(* IEC 61131-3 sources: plc-iiot-stack/src/POUs/Iiot/FB_MqttCommands, 19 files *)

(* ---- FB_MqttCommands.decl.st ---- *)
// Назначение: шлюз команд MQTT (data_schema 5): подписка <prefix>/+/cmd/+ (QoS 1), разбор подмножества JSON,
//             проверки по порядку раздела 5.1 (retained, invalid_payload, unsupported_version, topic_mismatch,
//             not_whitelisted, out_of_range, expired, duplicate, rate_limited) и ответ в
//             <prefix>/<device>/cmd_ack/<command>. Сообщение не своей станции или без читаемого cmd_id —
//             без ответа (udiDropped). Прошедшая команда — импульс xCmdValid и stCmd: вызывающий пишет её в
//             GVL_Hmi и вызывает Arm(); дальше ФБ ждёт, пока устройство увеличит uiCmdSeq (ok или
//             device_rejected по eCmdResult), иначе через tDeviceTimeout — timeout. Значения (SpeedSp) ФБ
//             устройства не квитирует: ok — сразу после записи. Одна команда в обработке за раз.
// Автор:      kr0nsch
// Версия:     0.1.0
// Документ:   docs/plc_mqtt.md, раздел «Команды»
FUNCTION_BLOCK FB_MqttCommands
VAR_INPUT
    xEnable : BOOL;
    itfClient : I_MqttClient;
    ltNow : LTIME;                                            // монотонное время (LTIME())
    uliTs_ms : ULINT;                                         // время UTC, мс: проверка ts и поле ts ответа
    sTopicPrefix : STRING(GVL_Const.IIOT_PREFIX_LEN);         // site/area/unit
    uiDevSeq : UINT;                                          // uiCmdSeq устройства команды в обработке
    iDevResult : INT;                                         // eCmdResult того же устройства
    tMaxAge : TIME := GVL_Const.CMD_MAX_AGE;
    tDeviceTimeout : TIME := GVL_Const.CMD_DEVICE_TIMEOUT;
    uiRateLimit : UINT := GVL_Const.CMD_RATE_LIMIT;           // не больше CMD_RATE_LIMIT
    tRateWindow : TIME := GVL_Const.CMD_RATE_WINDOW;
    uiMaxPerCycle : UINT := GVL_Const.CMD_MAX_PER_CYCLE;
END_VAR
VAR_IN_OUT
    aRules : ARRAY[*] OF ST_IiotCmdRule;                      // белый список
END_VAR
VAR_OUTPUT
    xCmdValid : BOOL;                                         // в этом вызове: записать stCmd в GVL_Hmi, затем Arm()
    stCmd : ST_IiotCmd;
    xPending : BOOL;                                          // ждём обработки устройством
    xSubscribed : BOOL;
    eLastReason : E_IiotCmdReason := E_IiotCmdReason.Ok;
    udiReceived : UDINT;
    udiAccepted : UDINT;                                      // ответов ok
    udiRejected : UDINT;                                      // ответов с отказом
    udiDropped : UDINT;                                       // без ответа: чужой топик, нет cmd_id
    udiAckFailed : UDINT;                                     // ответ не принят клиентом или не помещается
END_VAR
VAR
    fbParser : FB_JsonFlatParser;
    fbJson : FB_JsonBuilder;
    sFilter : STRING(GVL_Const.MQTT_TOPIC_LEN);
    sRxTopic : STRING(GVL_Const.MQTT_TOPIC_LEN);
    sRxPayload : STRING(GVL_Const.MQTT_CMD_PAYLOAD_LEN);
    xRxTruncated : BOOL;
    xRxRetained : BOOL;
    sAckTopic : STRING(GVL_Const.MQTT_TOPIC_LEN);
    // команда, на которую готовится ответ
    sTopicDevice : STRING(GVL_Const.IIOT_LEVEL_LEN);
    sTopicCommand : STRING(GVL_Const.IIOT_LEVEL_LEN);
    sCmdId : STRING(GVL_Const.JSON_STR_LEN);
    // повторы и частота
    aHistory : ARRAY[1..GVL_Const.CMD_HISTORY_LEN] OF STRING(GVL_Const.CMD_ID_LEN);
    uiHistoryNext : UINT := 1;
    aRateTimes : ARRAY[1..GVL_Const.CMD_RATE_LIMIT] OF LTIME;   // моменты последних прошедших команд
    uiRateNext : UINT := 1;
    uiRateCount : UINT;
    // обработка устройством
    xAwaitArm : BOOL;
    uiSeqArmed : UINT;
    ltPendingSince : LTIME;
    uiMsg : UINT;
END_VAR

(* ---- Arm.method.decl.st ---- *)
// Вызвать после записи stCmd в GVL_Hmi в том же цикле: uiSeqBefore — uiCmdSeq устройства до записи.
// Команды-значения (SpeedSp, SubstValue) отвечают ok сразу: ФБ устройства их не квитирует.
METHOD Arm
VAR_INPUT
    uiSeqBefore : UINT;
END_VAR

(* ---- Arm.method.impl.st ---- *)
IF NOT xAwaitArm THEN
    RETURN;
END_IF
xAwaitArm := FALSE;
IF F_IiotCmdKind(eCommand := stCmd.eCommand) = E_IiotCmdKind.Value THEN
    Finish(eReason := E_IiotCmdReason.Ok, iCmdResult := 0);
ELSE
    uiSeqArmed := uiSeqBefore;
    ltPendingSince := ltNow;
    xPending := TRUE;
END_IF

(* ---- Check.method.decl.st ---- *)
// Проверки шлюза по порядку data_schema 5.1, пункты 1–9; Ok — stCmd заполнена, момент учтён в частоте.
METHOD PRIVATE Check : E_IiotCmdReason
VAR_IN_OUT
    aRuleTable : ARRAY[*] OF ST_IiotCmdRule;
END_VAR
VAR
    sText : STRING(GVL_Const.JSON_STR_LEN);
    sKey : STRING(GVL_Const.JSON_KEY_LEN);
    iMajor : INT;
    uiIdx : UINT;
    lrTs : LREAL;
    lrValue : LREAL;
    lrMin : LREAL;
    lrMax : LREAL;
    xHasValue : BOOL;
    eCommand : E_IiotCommand;
    eKind : E_IiotCmdKind;
    diRule : DINT;
END_VAR

(* ---- Check.method.impl.st ---- *)
// 1. retained
IF xRxRetained THEN
    Check := E_IiotCmdReason.Retained;
    RETURN;
END_IF
// 2. состав и типы полей (command.schema.json; диапазон value — в п. 6)
Check := E_IiotCmdReason.InvalidPayload;
IF NOT fbParser.GetString(sKey := 'schema_version', sValue := sText) THEN
    RETURN;
END_IF
iMajor := F_IiotSchemaMajor(sVersion := sText);
IF iMajor < 0 THEN
    RETURN;
END_IF
FOR uiIdx := 1 TO fbParser.uiCount DO
    sKey := fbParser.KeyAt(uiIdx := uiIdx);
    IF sKey <> 'schema_version' AND sKey <> 'cmd_id' AND sKey <> 'ts' AND sKey <> 'origin' AND sKey <> 'command'
       AND sKey <> 'value' THEN
        RETURN;                     // лишнее поле: схема команды строгая
    END_IF
END_FOR
IF NOT fbParser.FieldIsInteger(sKey := 'ts') OR NOT fbParser.GetNumber(sKey := 'ts', lrValue := lrTs) THEN
    RETURN;
END_IF
IF lrTs < ULINT_TO_LREAL(GVL_Const.TS_MIN_MS) OR lrTs > ULINT_TO_LREAL(GVL_Const.TS_MAX_MS) THEN
    RETURN;
END_IF
IF NOT fbParser.GetString(sKey := 'origin', sValue := sText) THEN
    RETURN;
END_IF
IF NOT F_IiotIsPrintable(sText := sText, iMaxLen := UINT_TO_INT(GVL_Const.CMD_ORIGIN_LEN)) THEN
    RETURN;
END_IF
IF NOT fbParser.GetString(sKey := 'command', sValue := sText) THEN
    RETURN;
END_IF
eCommand := F_IiotCmdFromString(sCommand := sText);
IF eCommand = E_IiotCommand.None THEN
    RETURN;
END_IF
eKind := F_IiotCmdKind(eCommand := eCommand);
xHasValue := fbParser.FieldType(sKey := 'value') <> E_JsonType.Missing;
IF xHasValue AND NOT fbParser.GetNumber(sKey := 'value', lrValue := lrValue) THEN
    RETURN;                         // value не число
END_IF
IF eKind = E_IiotCmdKind.Pulse AND xHasValue THEN
    RETURN;                         // value у импульсной команды
END_IF
IF eKind <> E_IiotCmdKind.Pulse AND NOT xHasValue THEN
    RETURN;                         // нет value
END_IF
IF eKind = E_IiotCmdKind.Mask
   AND (NOT fbParser.FieldIsInteger(sKey := 'value') OR lrValue < 0.0 OR lrValue > GVL_Const.CMD_MASK_MAX) THEN
    RETURN;                         // маска: целое 0..65535
END_IF
// 3. мажорная версия
IF iMajor <> UINT_TO_INT(GVL_Const.IIOT_SCHEMA_MAJOR) THEN
    Check := E_IiotCmdReason.UnsupportedVersion;
    RETURN;
END_IF
// 4. команда в теле и в топике
IF sText <> sTopicCommand THEN
    Check := E_IiotCmdReason.TopicMismatch;
    RETURN;
END_IF
// 5. белый список
diRule := FindRule(aRuleTable := aRuleTable, eCommandIn := eCommand);
IF diRule < LOWER_BOUND(aRuleTable, 1) THEN
    Check := E_IiotCmdReason.NotWhitelisted;
    RETURN;
END_IF
// 6. диапазон значения
IF xHasValue THEN
    IF aRuleTable[diRule].xRange THEN
        lrMin := REAL_TO_LREAL(aRuleTable[diRule].rMin);
        lrMax := REAL_TO_LREAL(aRuleTable[diRule].rMax);
    ELSE
        lrMin := -GVL_Const.REAL_ABS_MAX;
        lrMax := GVL_Const.REAL_ABS_MAX;
    END_IF
    IF eCommand = E_IiotCommand.SpeedSp THEN       // схема: 0..100 % независимо от белого списка
        lrMin := MAX(lrMin, GVL_Const.SPEED_SP_MIN_PCT);
        lrMax := MIN(lrMax, GVL_Const.SPEED_SP_MAX_PCT);
    END_IF
    IF lrValue < lrMin OR lrValue > lrMax THEN
        Check := E_IiotCmdReason.OutOfRange;
        RETURN;
    END_IF
END_IF
// 7. возраст ts (часы ПЛК должны быть установлены)
IF NOT F_IiotClockValid(uliTs_ms := uliTs_ms)
   OR ABS(ULINT_TO_LREAL(uliTs_ms) - lrTs) > ULINT_TO_LREAL(TIME_TO_ULINT(tMaxAge)) THEN
    Check := E_IiotCmdReason.Expired;
    RETURN;
END_IF
// 8. повтор cmd_id
IF IsDuplicate() THEN
    Check := E_IiotCmdReason.Duplicate;
    RETURN;
END_IF
// 9. частота
IF NOT RateAllows() THEN
    Check := E_IiotCmdReason.RateLimited;
    RETURN;
END_IF
stCmd.diRule := diRule;
stCmd.sDevice := sTopicDevice;
stCmd.sCommand := sTopicCommand;
stCmd.eCommand := eCommand;
stCmd.rValue := LREAL_TO_REAL(lrValue);
stCmd.sCmdId := sCmdId;
Check := E_IiotCmdReason.Ok;

(* ---- FB_MqttCommands.impl.st ---- *)
xCmdValid := FALSE;
IF NOT xEnable OR itfClient = 0 THEN
    xSubscribed := FALSE;
    xPending := FALSE;
    xAwaitArm := FALSE;
    RETURN;
END_IF
IF NOT itfClient.IsConnected() THEN
    xSubscribed := FALSE;     // после подключения — подписка заново (сессия может быть чистой)
    RETURN;
END_IF
IF NOT xSubscribed THEN
    sFilter := CONCAT(sTopicPrefix, GVL_Const.TOPIC_CMD_FILTER_SUFFIX);
    xSubscribed := itfClient.Subscribe(sTopicFilter := sFilter, eQos := E_MqttQos.AtLeastOnce);
    IF NOT xSubscribed THEN
        RETURN;
    END_IF
END_IF

// Команда прошла проверки в прошлом вызове, но Arm() не вызван: до устройства она не дошла
IF xAwaitArm THEN
    xAwaitArm := FALSE;
    Finish(eReason := E_IiotCmdReason.Timeout, iCmdResult := 0);
END_IF
// Команда в обработке устройством
IF xPending THEN
    IF uiDevSeq <> uiSeqArmed AND iDevResult >= GVL_Const.CMD_RESULT_ACCEPTED
       AND iDevResult <= GVL_Const.CMD_RESULT_LAST THEN
        xPending := FALSE;
        IF iDevResult = GVL_Const.CMD_RESULT_ACCEPTED THEN
            Finish(eReason := E_IiotCmdReason.Ok, iCmdResult := iDevResult);
        ELSE
            Finish(eReason := E_IiotCmdReason.DeviceRejected, iCmdResult := iDevResult);
        END_IF
    ELSIF ltNow < ltPendingSince THEN
        ltPendingSince := ltNow;
    ELSIF (ltNow - ltPendingSince) >= TIME_TO_LTIME(tDeviceTimeout) THEN
        xPending := FALSE;
        Finish(eReason := E_IiotCmdReason.Timeout, iCmdResult := 0);
    END_IF
    IF xPending THEN
        RETURN;
    END_IF
END_IF

FOR uiMsg := 1 TO MAX(uiMaxPerCycle, 1) DO
    IF xCmdValid THEN
        EXIT;
    END_IF
    IF NOT itfClient.Receive(sTopic := sRxTopic, sPayload := sRxPayload, xTruncated => xRxTruncated,
                             xRetained => xRxRetained) THEN
        EXIT;
    END_IF
    udiReceived := udiReceived + 1;
    HandleMessage(aRuleTable := aRules);
END_FOR

(* ---- FindRule.method.decl.st ---- *)
// Строка белого списка для (sTopicDevice, eCommandIn); нет — LOWER_BOUND - 1.
METHOD PRIVATE FindRule : DINT
VAR_IN_OUT
    aRuleTable : ARRAY[*] OF ST_IiotCmdRule;
END_VAR
VAR_INPUT
    eCommandIn : E_IiotCommand;
END_VAR
VAR
    diIdx : DINT;
END_VAR

(* ---- FindRule.method.impl.st ---- *)
FindRule := LOWER_BOUND(aRuleTable, 1) - 1;
FOR diIdx := LOWER_BOUND(aRuleTable, 1) TO UPPER_BOUND(aRuleTable, 1) DO
    IF aRuleTable[diIdx].eCommand = eCommandIn AND aRuleTable[diIdx].sDevice = sTopicDevice THEN
        FindRule := diIdx;
        RETURN;
    END_IF
END_FOR

(* ---- Finish.method.decl.st ---- *)
// Ответ в <prefix>/<sTopicDevice>/cmd_ack/<sTopicCommand>: schema_version, cmd_id, ts, command, result, reason
// и cmd_result (device_rejected). Счётчики принятых и отклонённых команд.
METHOD PRIVATE Finish
VAR_INPUT
    eReason : E_IiotCmdReason;
    iCmdResult : INT;             // E_CmdResult устройства; 0 — нет
END_VAR
VAR
    sResultText : STRING(GVL_Const.IIOT_TEXT_LEN);
    sPath : STRING(GVL_Const.MQTT_TOPIC_LEN);
END_VAR

(* ---- Finish.method.impl.st ---- *)
eLastReason := eReason;
IF eReason = E_IiotCmdReason.Ok THEN
    udiAccepted := udiAccepted + 1;
ELSE
    udiRejected := udiRejected + 1;
END_IF
sPath := CONCAT(CONCAT(sTopicDevice, GVL_Const.TOPIC_SEPARATOR), GVL_Const.TOPIC_ACK_LEVEL);
sPath := CONCAT(CONCAT(sPath, GVL_Const.TOPIC_SEPARATOR), sTopicCommand);
sAckTopic := F_IiotTopic(sPrefix := sTopicPrefix, sPath := sPath);
fbJson.Begin();
fbJson.AddString(sKey := 'schema_version', sValue := GVL_Const.IIOT_SCHEMA_VERSION);
fbJson.AddString(sKey := 'cmd_id', sValue := sCmdId);
fbJson.AddInt(sKey := 'ts', liValue := ULINT_TO_LINT(uliTs_ms));
fbJson.AddString(sKey := 'command', sValue := sTopicCommand);
IF eReason = E_IiotCmdReason.Ok THEN
    fbJson.AddString(sKey := 'result', sValue := 'accepted');
ELSE
    fbJson.AddString(sKey := 'result', sValue := 'rejected');
END_IF
fbJson.AddString(sKey := 'reason', sValue := F_IiotCmdReasonText(eReason := eReason));
sResultText := F_IiotCmdResultText(iResult := iCmdResult);
IF eReason = E_IiotCmdReason.DeviceRejected AND LEN(sResultText) > 0 THEN
    fbJson.AddString(sKey := 'cmd_result', sValue := sResultText);
END_IF
IF NOT fbJson.Finish() OR LEN(sAckTopic) = 0 THEN
    udiAckFailed := udiAckFailed + 1;
ELSIF NOT itfClient.Publish(sTopic := sAckTopic, eQos := E_MqttQos.AtLeastOnce, xRetain := FALSE,
                            sPayload := fbJson.sJson) THEN
    udiAckFailed := udiAckFailed + 1;
END_IF

(* ---- HandleMessage.method.decl.st ---- *)
// Разбор принятого сообщения: без ответа (чужой топик, нет cmd_id), отказ с ответом или команда в stCmd.
METHOD PRIVATE HandleMessage
VAR_IN_OUT
    aRuleTable : ARRAY[*] OF ST_IiotCmdRule;
END_VAR
VAR
    eReason : E_IiotCmdReason;
END_VAR

(* ---- HandleMessage.method.impl.st ---- *)
sCmdId := '';
IF NOT SplitTopic() THEN
    udiDropped := udiDropped + 1;      // не команда своей станции — отвечать некуда
    RETURN;
END_IF
IF xRxTruncated OR NOT fbParser.Parse(sJson := sRxPayload) THEN
    udiDropped := udiDropped + 1;      // не JSON-объект: cmd_id не прочитать
    RETURN;
END_IF
IF NOT fbParser.GetString(sKey := 'cmd_id', sValue := sCmdId) OR NOT F_IiotIsCmdId(sText := sCmdId) THEN
    sCmdId := '';
    udiDropped := udiDropped + 1;
    RETURN;
END_IF
eReason := Check(aRuleTable := aRuleTable);
IF eReason <> E_IiotCmdReason.Duplicate THEN
    Remember();
END_IF
IF eReason = E_IiotCmdReason.Ok THEN
    xCmdValid := TRUE;
    xAwaitArm := TRUE;
ELSE
    Finish(eReason := eReason, iCmdResult := 0);
END_IF

(* ---- IsDuplicate.method.decl.st ---- *)
// cmd_id текущей команды встречался среди последних CMD_HISTORY_LEN.
METHOD PRIVATE IsDuplicate : BOOL
VAR
    uiIdx : UINT;
END_VAR

(* ---- IsDuplicate.method.impl.st ---- *)
FOR uiIdx := 1 TO GVL_Const.CMD_HISTORY_LEN DO
    IF LEN(aHistory[uiIdx]) > 0 AND aHistory[uiIdx] = sCmdId THEN
        IsDuplicate := TRUE;
        RETURN;
    END_IF
END_FOR

(* ---- RateAllows.method.decl.st ---- *)
// Частота: не больше uiRateLimit прошедших команд за tRateWindow. TRUE — команда разрешена и учтена.
METHOD PRIVATE RateAllows : BOOL
VAR
    uiLimit : UINT;
END_VAR

(* ---- RateAllows.method.impl.st ---- *)
uiLimit := MIN(MAX(uiRateLimit, 1), GVL_Const.CMD_RATE_LIMIT);
IF uiRateNext < 1 OR uiRateNext > uiLimit THEN
    uiRateNext := 1;
END_IF
// в кольце из uiLimit моментов следующая позиция — самая старая из последних uiLimit команд
IF uiRateCount >= uiLimit AND_THEN ltNow >= aRateTimes[uiRateNext]
   AND_THEN (ltNow - aRateTimes[uiRateNext]) <= TIME_TO_LTIME(tRateWindow) THEN
    RETURN;
END_IF
aRateTimes[uiRateNext] := ltNow;
uiRateNext := uiRateNext + 1;
IF uiRateNext > uiLimit THEN
    uiRateNext := 1;
END_IF
IF uiRateCount < uiLimit THEN
    uiRateCount := uiRateCount + 1;
END_IF
RateAllows := TRUE;

(* ---- Remember.method.impl.st ---- *)
IF uiHistoryNext < 1 OR uiHistoryNext > GVL_Const.CMD_HISTORY_LEN THEN
    uiHistoryNext := 1;
END_IF
aHistory[uiHistoryNext] := sCmdId;
uiHistoryNext := uiHistoryNext + 1;

(* ---- SplitTopic.method.decl.st ---- *)
// Разобрать sRxTopic вида <prefix>/<DEVICE>/cmd/<Command> в sTopicDevice и sTopicCommand. FALSE — топик не
// своей станции или уровни не по шаблонам ([A-Z][A-Z0-9_]{0,15} и [A-Za-z][A-Za-z0-9_]{0,31}).
METHOD PRIVATE SplitTopic : BOOL
VAR
    iPrefixLen : INT;
    sRest : STRING(GVL_Const.MQTT_TOPIC_LEN);
    sTail : STRING(GVL_Const.MQTT_TOPIC_LEN);
    iSlash : INT;
END_VAR

(* ---- SplitTopic.method.impl.st ---- *)
sTopicDevice := '';
sTopicCommand := '';
iPrefixLen := LEN(sTopicPrefix);
IF iPrefixLen = 0 OR LEN(sRxTopic) <= iPrefixLen + 1 THEN
    RETURN;
END_IF
IF LEFT(sRxTopic, iPrefixLen) <> sTopicPrefix OR MID(sRxTopic, 1, iPrefixLen + 1) <> GVL_Const.TOPIC_SEPARATOR THEN
    RETURN;
END_IF
sRest := RIGHT(sRxTopic, LEN(sRxTopic) - iPrefixLen - 1);
// <DEVICE>
iSlash := FIND(sRest, GVL_Const.TOPIC_SEPARATOR);
IF iSlash <= 1 OR iSlash - 1 > UINT_TO_INT(GVL_Const.IIOT_DEVICE_LEN) THEN
    RETURN;
END_IF
sTopicDevice := LEFT(sRest, iSlash - 1);
sTail := RIGHT(sRest, LEN(sRest) - iSlash);
// cmd
iSlash := FIND(sTail, GVL_Const.TOPIC_SEPARATOR);
IF iSlash <= 1 OR LEFT(sTail, iSlash - 1) <> GVL_Const.TOPIC_CMD_LEVEL THEN
    sTopicDevice := '';
    RETURN;
END_IF
// <Command>
IF LEN(sTail) - iSlash > UINT_TO_INT(GVL_Const.IIOT_LEVEL_LEN) THEN
    sTopicDevice := '';
    RETURN;
END_IF
sTopicCommand := RIGHT(sTail, LEN(sTail) - iSlash);
IF NOT F_IiotIsName(sText := sTopicDevice, iMaxLen := UINT_TO_INT(GVL_Const.IIOT_DEVICE_LEN), xUpperOnly := TRUE)
   OR NOT F_IiotIsName(sText := sTopicCommand, iMaxLen := UINT_TO_INT(GVL_Const.IIOT_LEVEL_LEN),
                       xUpperOnly := FALSE) THEN
    sTopicDevice := '';
    sTopicCommand := '';
    RETURN;
END_IF
SplitTopic := TRUE;
